// TIA Portal V19 export
DATA_BLOCK "START_DB"   // DB19
// stored: InstanceOfName START, InstanceOfType FB
"START"
   // VAR_INPUT
   //    RUNNING : Bool;
   // END_VAR
   // VAR_OUTPUT
   //    START_CMD : Bool;
   //    STOP_CMD : Bool;
   // END_VAR
   // VAR_IN_OUT
   //    "START/STOP" : Bool;
   // END_VAR
   // VAR
   //    START_PLS : Bool;
   //    IEC_Timer_0_Instance { S7_SetPoint := 'True'} : TOF_TIME;
   //    STOP_PLS : Bool;
   //    IEC_Timer_0_Instance_1 { S7_SetPoint := 'True'} : TOF_TIME;
   //    RUNNING_PLS : Bool;
   //    "HEAT/COOL_Instance" { S7_SetPoint := 'True'} : "HEAT/COOL";
   // END_VAR
BEGIN
END_DATA_BLOCK
